// TIA Portal V20 export
// export: Created 2026-10-12T05:42:29.8554295Z, ExportSetting WithDefaults, DisplayName Totally Integrated Automation Portal, DisplayVersion V20, DisplayName TIA Portal Openness, DisplayVersion V20, DisplayName TIA Portal Teamcenter Gateway, DisplayVersion V20, DisplayName TIA Portal Version Control Interface, DisplayVersion V20, DisplayName SINAMICS Startdrive Advanced, DisplayVersion V20 SP1 Update 2, DisplayName SINAMICS Startdrive G110M, G120, G120C, G120D, G120P, G115D, DisplayVersion V20 SP1 Update 2, DisplayName SINAMICS Startdrive G130, G150, S120, S150, SINAMICS MV, G220, S200, S210, DisplayVersion V20 SP1 Update 2, DisplayName STEP 7 Professional, DisplayVersion V20, DisplayName STEP 7 Safety, DisplayVersion V20, DisplayName WinCC Basic/Comfort/Advanced, DisplayVersion V20, DisplayName WinCC Professional, DisplayVersion V20, DisplayName WinCC Unified, DisplayVersion V20
FUNCTION "FRK_AccessUsersCrc" : DWord   // FC50, SCL
{ S7_Optimized_Access := 'TRUE' }
VERSION : 0.1
// stored: AutoNumber true, IsIECCheckEnabled false, SetENOAutomatically false, UDAEnableTagReadback false
   VAR_TEMP
      Work : DWord;
      Slot : Int;
      Index : Int;
      Size : Int;
   END_VAR
BEGIN

   #Work := "FRK_AccessCrcNumber"(Previous := DWORD#16#FFFFFFFF, Value := UINT_TO_UDINT("FRK_LocalUsers".SchemaVersion));
   #Work := "FRK_AccessCrcNumber"(Previous := #Work, Value := "FRK_LocalUsers".Generation);
   #Work := "FRK_AccessCrcNumber"(Previous := #Work, Value := DINT_TO_UDINT("FRK_LocalUsers".Count));
   // Unused rows are included: an altered dormant credential is not ignored.
   FOR #Slot := 1 TO 16 DO
       #Size := LEN("FRK_LocalUsers".Rows[#Slot].User);
       #Work := "FRK_AccessCrcNumber"(Previous := #Work, Value := INT_TO_UDINT(#Size));
       FOR #Index := 1 TO #Size DO
           #Work := "FRK_AccessCrcByte"(Previous := #Work, Value := CHAR_TO_BYTE("FRK_LocalUsers".Rows[#Slot].User[#Index]));
       END_FOR;
       #Work := "FRK_AccessCrcNumber"(Previous := #Work, Value := DINT_TO_UDINT("FRK_LocalUsers".Rows[#Slot].Level));
       FOR #Index := 0 TO 15 DO
           #Work := "FRK_AccessCrcByte"(Previous := #Work, Value := "FRK_LocalUsers".Rows[#Slot].Salt[#Index]);
       END_FOR;
       FOR #Index := 0 TO 31 DO
           #Work := "FRK_AccessCrcByte"(Previous := #Work, Value := "FRK_LocalUsers".Rows[#Slot].PinHash[#Index]);
       END_FOR;
   END_FOR;
   #FRK_AccessUsersCrc := NOT #Work;
END_FUNCTION
